Fanuc KAREL source: KT00537.KL

PROGRAM KT00537
%NOLOCKGROUP
VAR
  P1: JOINTPOS
  P2: POSITION
  OUT: JOINTPOS
BEGIN
  OUT = P1 : P2
END KT00537
